FUNCTION F_UpsSignedWord : REAL
VAR_INPUT i_wRaw : WORD; END_VAR

IF i_wRaw >= 16#8000 THEN
	F_UpsSignedWord := DINT_TO_REAL(WORD_TO_DINT(i_wRaw) - 65536);
ELSE
	F_UpsSignedWord := WORD_TO_REAL(i_wRaw);
END_IF

END_FUNCTION

(* stored: Version 1.1.0.1, ProductVersion 3.1.4024.15
   POU F_UpsSignedWord: Id {3332eb93-bedd-4662-9d1c-253a8424a0dc} *)
